// TIA Portal V19 export
// export: Created 2026-10-15T10:10:34.7901659Z, ExportSetting WithDefaults, DisplayName Totally Integrated Automation Portal, DisplayVersion V19, DisplayName TIA Portal Openness, DisplayVersion V19, DisplayName TIA Portal Version Control Interface, DisplayVersion V19, DisplayName STEP 7 Professional, DisplayVersion V19, DisplayName STEP 7 Safety, DisplayVersion V19, DisplayName WinCC Basic/Comfort/Advanced, DisplayVersion V19, DisplayName WinCC Unified, DisplayVersion V19
FUNCTION "ROLL_DecodeBCD" : Int   // FC4, SCL
{ S7_Optimized_Access := 'TRUE' }
VERSION : 0.1
// stored: AutoNumber true, IsIECCheckEnabled false, SetENOAutomatically false, UDAEnableTagReadback false
   VAR_INPUT
      Value : Word;
   END_VAR
   VAR_TEMP
      hundreds : Int;
      tens : Int;
      units : Int;
   END_VAR
BEGIN

   #hundreds := WORD_TO_INT(SHR(IN := #Value AND W#16#0F00, N := 8));
   #tens := WORD_TO_INT(SHR(IN := #Value AND W#16#00F0, N := 4));
   #units := WORD_TO_INT(#Value AND W#16#000F);
   IF (#hundreds > 9) OR (#tens > 9) OR (#units > 9) THEN
       "ROLL_IO".ConversionFault := TRUE;
       #ROLL_DecodeBCD := -1;
   ELSE
       #ROLL_DecodeBCD := #hundreds * 100 + #tens * 10 + #units;
   END_IF;
END_FUNCTION
